Staubli VAL3: utAppearance.dtx

public string sBackgroundColour
public bool bVisibility
